Omron CX-Programmer project NewProject (CX-Programmer 9.81)

# PLC masodik: CJ2M CPU32
I/O table (CPU CJ2M-CPU32): rack 0 slot 11 CJ2M-EIP21

## Global symbols (name address type ; comment)
At_entry 2.00 BOOL  ; At entry
At_front 2.06 BOOL  ; At front
At_left_entry 2.08 BOOL  ; At left entry
At_left_exit 2.10 BOOL  ; At left exit
At_load_position 2.04 BOOL  ; At load position
At_right_entry 2.07 BOOL  ; At right entry
At_right_exit 2.09 BOOL  ; At right exit
At_turntable_entry 2.03 BOOL  ; At turntable entry
At_unload_position 2.05 BOOL  ; At unload position
Emergency_stop 2.14 BOOL  ; Emergency stop
Entry_conveyor 3.01 BOOL  ; Entry conveyor
Feeder_conveyor 3.00 BOOL  ; Feeder conveyor
Green_indicator 3.07 BOOL  ; Green indicator
High_box 2.02 BOOL  ; High box
Left_conveyor 3.05 BOOL  ; Left conveyor
Load 3.02 BOOL  ; Load
Low_box 2.01 BOOL  ; Low box
Red_indicator 3.09 BOOL  ; Red indicator
Reset 2.12 BOOL  ; Reset
Reset_light 3.11 BOOL  ; Reset light
Right_conveyor 3.06 BOOL  ; Right conveyor
Start 2.11 BOOL  ; Start
Start_light 3.10 BOOL  ; Start light
Stop 2.13 BOOL  ; Stop
Stop_light 3.12 BOOL  ; Stop light
Turn 3.04 BOOL  ; Turn
Unload 3.03 BOOL  ; Unload
Yellow_indicator 3.08 BOOL  ; Yellow indicator
a_num W350 UINT
b_num W351 UINT
dest W352 UINT
next_prod W200 UINT

## Program NewProgram2 (cyclic task 0)
Local symbols
enable W0.00 BOOL
left_counter W4 UINT
right_counter W5 UINT
stack_length W6 UINT
stack_light UINT
stack_null W0.04 BOOL
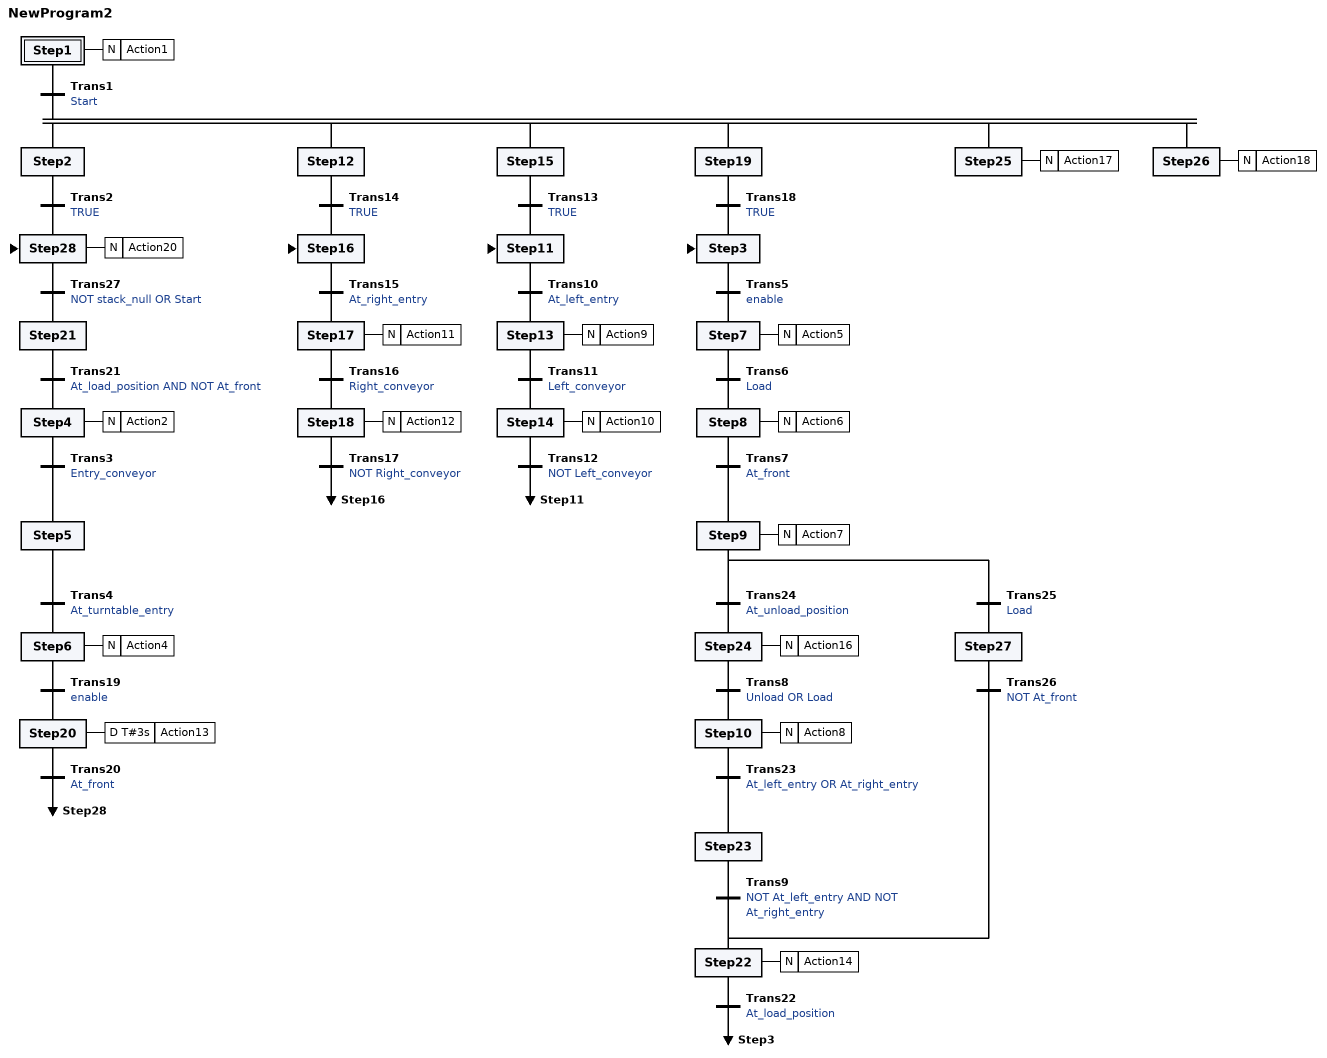
INITIAL_STEP Step1 :
Action1(N) ;
END_STEP
TRANSITION Trans1 FROM Step1 TO (Step2,Step12,Step15,Step19,Step25,Step26)
 := Start;
END_TRANSITION
STEP Step2 :
END_STEP
STEP Step3 :
END_STEP
TRANSITION Trans2 FROM Step2 TO Step28
 := TRUE;
END_TRANSITION
STEP Step4 :
Action2(N) ;
END_STEP
TRANSITION Trans3 FROM Step4 TO Step5
 := Entry_conveyor;
END_TRANSITION
STEP Step5 :
END_STEP
TRANSITION Trans4 FROM Step5 TO Step6
 := At_turntable_entry;
END_TRANSITION
STEP Step6 :
Action4(N) ;
END_STEP
TRANSITION Trans5 FROM Step3 TO Step7
 := enable;
END_TRANSITION
STEP Step7 :
Action5(N) ;
END_STEP
TRANSITION Trans6 FROM Step7 TO Step8
 := Load;
END_TRANSITION
STEP Step8 :
Action6(N) ;
END_STEP
TRANSITION Trans7 FROM Step8 TO Step9
 := At_front;
END_TRANSITION
STEP Step9 :
Action7(N) ;
END_STEP
TRANSITION Trans8 FROM Step24 TO Step10
 := Unload OR Load;
END_TRANSITION
STEP Step11 :
END_STEP
STEP Step12 :
END_STEP
TRANSITION Trans10 FROM Step11 TO Step13
 := At_left_entry;
END_TRANSITION
STEP Step13 :
Action9(N) ;
END_STEP
TRANSITION Trans11 FROM Step13 TO Step14
 := Left_conveyor;
END_TRANSITION
STEP Step14 :
Action10(N) ;
END_STEP
STEP Step10 :
Action8(N) ;
END_STEP
TRANSITION Trans9 FROM Step23 TO Step22
 := NOT At_left_entry AND NOT At_right_entry;
END_TRANSITION
TRANSITION Trans12 FROM Step14 TO Step11
 := NOT Left_conveyor;
END_TRANSITION
STEP Step15 :
END_STEP
TRANSITION Trans13 FROM Step15 TO Step11
 := TRUE;
END_TRANSITION
TRANSITION Trans14 FROM Step12 TO Step16
 := TRUE;
END_TRANSITION
STEP Step16 :
END_STEP
TRANSITION Trans15 FROM Step16 TO Step17
 := At_right_entry;
END_TRANSITION
STEP Step17 :
Action11(N) ;
END_STEP
TRANSITION Trans16 FROM Step17 TO Step18
 := Right_conveyor;
END_TRANSITION
STEP Step18 :
Action12(N) ;
END_STEP
TRANSITION Trans17 FROM Step18 TO Step16
 := NOT Right_conveyor;
END_TRANSITION
STEP Step19 :
END_STEP
TRANSITION Trans18 FROM Step19 TO Step3
 := TRUE;
END_TRANSITION
TRANSITION Trans19 FROM Step6 TO Step20
 := enable;
END_TRANSITION
STEP Step20 :
Action13(D,T#3s) ;
END_STEP
TRANSITION Trans20 FROM Step20 TO Step28
 := At_front;
END_TRANSITION
STEP Step21 :
END_STEP
TRANSITION Trans21 FROM Step21 TO Step4
 := At_load_position AND NOT At_front;
END_TRANSITION
STEP Step22 :
Action14(N) ;
END_STEP
TRANSITION Trans22 FROM Step22 TO Step3
 := At_load_position;
END_TRANSITION
TRANSITION Trans23 FROM Step10 TO Step23
 := At_left_entry OR At_right_entry;
END_TRANSITION
STEP Step23 :
END_STEP
STEP Step24 :
Action16(N) ;
END_STEP
STEP Step25 :
Action17(N) ;
END_STEP
STEP Step26 :
Action18(N) ;
END_STEP
TRANSITION Trans24 (PRIORITY := 1) FROM Step9 TO Step24
 := At_unload_position;
END_TRANSITION
TRANSITION Trans25 (PRIORITY := 2) FROM Step9 TO Step27
 := Load;
END_TRANSITION
STEP Step27 :
END_STEP
TRANSITION Trans26 FROM Step27 TO Step22
 := NOT At_front;
END_TRANSITION
STEP Step28 :
Action20(N) ;
END_STEP
TRANSITION Trans27 FROM Step28 TO Step21
 := NOT stack_null OR Start;
END_TRANSITION

### Action Action1

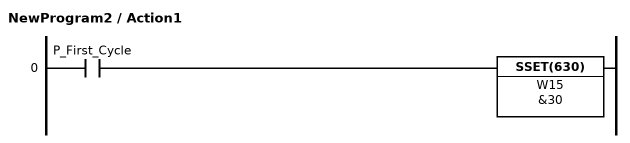
; rung 0
LD P_First_Cycle
SSET(630) W15 &30

### Action Action2

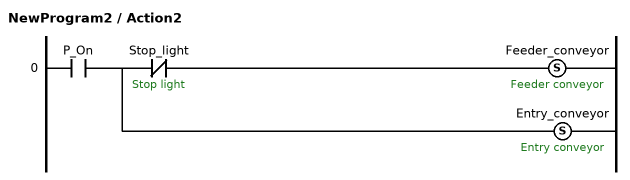
; rung 0
LD P_On
OUT TR0
ANDNOT Stop_light  ; Stop light
SET Feeder_conveyor  ; Feeder conveyor
LD TR0
SET Entry_conveyor  ; Entry conveyor

### Action Action3

### Action Action4

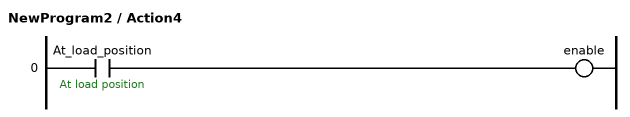
; rung 0
LD At_load_position  ; At load position
OUT enable

### Action Action5

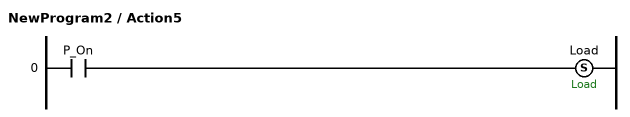
; rung 0
LD P_On
SET Load  ; Load

### Action Action6

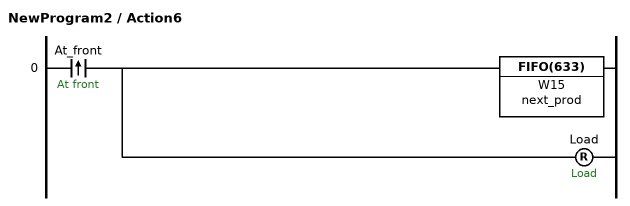
; rung 0
@LD At_front  ; At front
FIFO(633) W15 next_prod
RSET Load  ; Load

### Action Action7

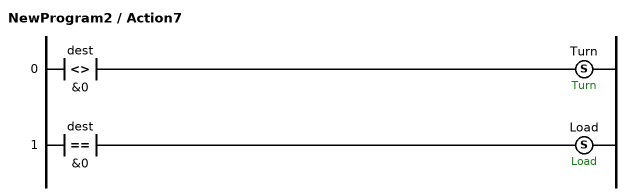
; rung 0
LD<>(305) dest &0
SET Turn  ; Turn
; rung 1
LD=(300) dest &0
SET Load  ; Load

### Action Action8

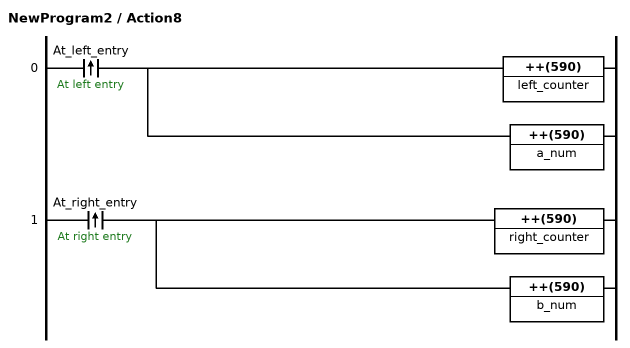
; rung 0
@LD At_left_entry  ; At left entry
++(590) left_counter
++(590) a_num
; rung 1
@LD At_right_entry  ; At right entry
++(590) right_counter
++(590) b_num

### Action Action9

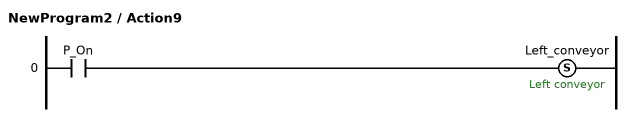
; rung 0
LD P_On
SET Left_conveyor  ; Left conveyor

### Action Action10

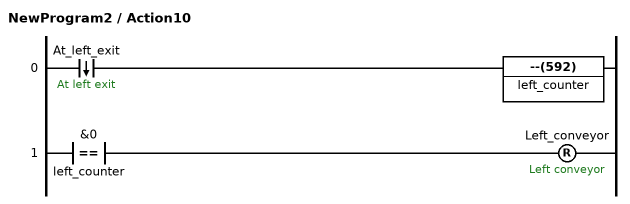
; rung 0
%LD At_left_exit  ; At left exit
--(592) left_counter
; rung 1
LD=(300) &0 left_counter
RSET Left_conveyor  ; Left conveyor

### Action Action11

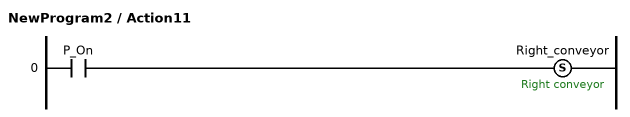
; rung 0
LD P_On
SET Right_conveyor  ; Right conveyor

### Action Action12

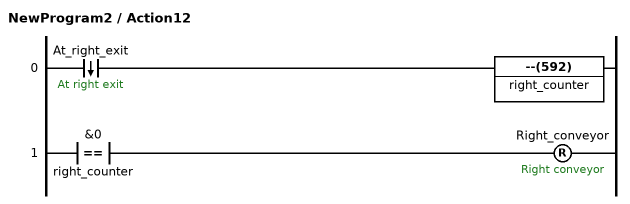
; rung 0
%LD At_right_exit  ; At right exit
--(592) right_counter
; rung 1
LD=(300) &0 right_counter
RSET Right_conveyor  ; Right conveyor

### Action Action13

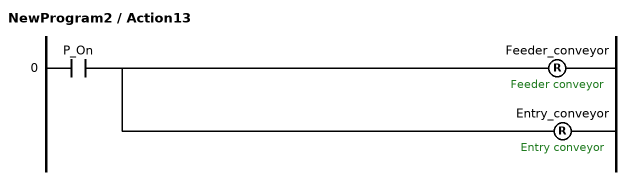
; rung 0
LD P_On
RSET Feeder_conveyor  ; Feeder conveyor
RSET Entry_conveyor  ; Entry conveyor

### Action Action14

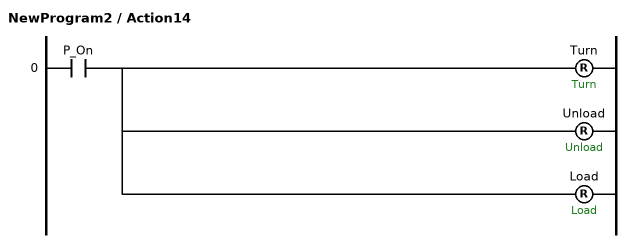
; rung 0
LD P_On
RSET Turn  ; Turn
RSET Unload  ; Unload
RSET Load  ; Load

### Action Action15

### Action Action16

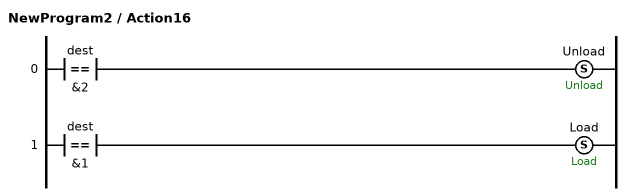
; rung 0
LD=(300) dest &2
SET Unload  ; Unload
; rung 1
LD=(300) dest &1
SET Load  ; Load

### Action Action17

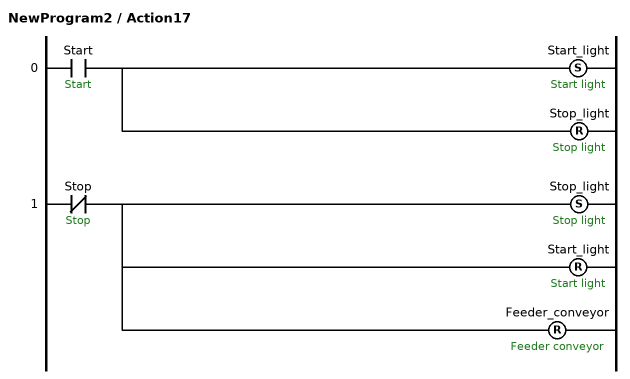
; rung 0
LD Start  ; Start
SET Start_light  ; Start light
RSET Stop_light  ; Stop light
; rung 1
LDNOT Stop  ; Stop
SET Stop_light  ; Stop light
RSET Start_light  ; Start light
RSET Feeder_conveyor  ; Feeder conveyor

### Action Action18

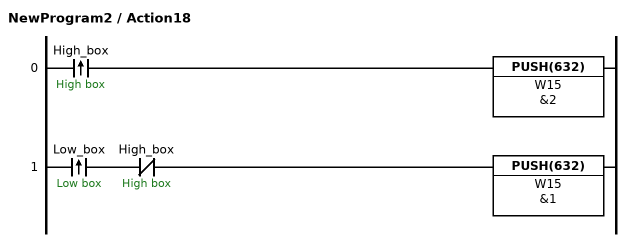
; rung 0
@LD High_box  ; High box
PUSH(632) W15 &2
; rung 1
@LD Low_box  ; Low box
ANDNOT High_box  ; High box
PUSH(632) W15 &1

### Action Action19

### Action Action20

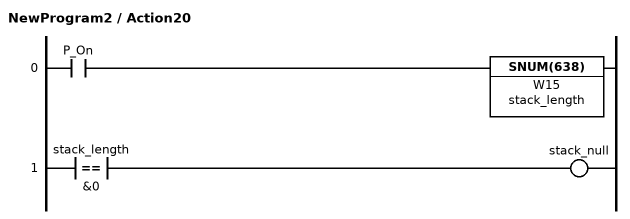
; rung 0
LD P_On
SNUM(638) W15 stack_length
; rung 1
LD=(300) stack_length &0
OUT stack_null

## Program NewProgram3 (cyclic task 1)
Local symbols
a_array W500 UINT[4]
a_comp W0.01 BOOL
b_array W400 UINT[6]
b_comp W0.02 BOOL
IF P_First_Cycle THEN
	a_num := 0;
	b_num := 0;
	a_comp := FALSE;
	b_comp := FALSE;
	
	a_array[0] := 1;
	a_array[1] := 2;
	a_array[2] := 1;
	a_array[3] := 2;
	
	b_array[0] := 1;
	b_array[1] := 1;
	b_array[2] := 1;
	b_array[3] := 2;
	b_array[4] := 2;
	b_array[5] := 2;
END_IF;

IF a_comp AND b_comp THEN
	dest := 0;
ELSIF a_comp AND b_array[b_num] = next_prod THEN
	dest := 2;
ELSIF b_comp AND a_array[a_num] = next_prod THEN
	dest := 1;
ELSIF next_prod = 1 THEN
	IF a_array[a_num] <> 1 AND b_array[b_num] <> 1 THEN
		dest := 0;
	ELSIF a_array[a_num] = 1 AND b_array[b_num] <> 1 THEN
		dest := 1;
	ELSIF a_array[a_num] <> 1 AND b_array[b_num] = 1 THEN
		dest := 2;
	ELSIF a_array[a_num] = 1 AND b_array[b_num] = 1 THEN
		IF a_num > b_num THEN
			dest := 2;
		ELSIF a_num < b_num THEN
			dest := 1;
		ELSE
			dest := 1;
		END_IF;
	END_IF;
ELSIF next_prod = 2 THEN
	IF a_array[a_num] <> 2 AND b_array[b_num] <> 2 THEN
		dest := 0;
	ELSIF a_array[a_num] = 2 AND b_array[b_num] <> 2 THEN
		dest := 1;
	ELSIF a_array[a_num] <> 2 AND b_array[b_num] = 2 THEN
		dest := 2;
	ELSIF a_array[a_num] = 2 AND b_array[b_num] = 2 THEN
		IF a_num > b_num THEN
			dest := 2;
		ELSIF a_num < b_num THEN
			dest := 1;
		ELSE
			dest := 1;
		END_IF;
	END_IF;
END_IF;

## Program NewProgram1 (cyclic task 2)
Local symbols
Emergency_light BOOL
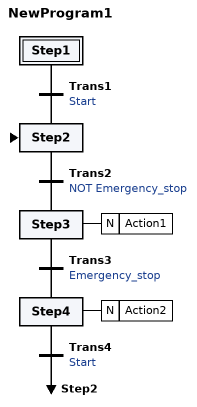
INITIAL_STEP Step1 :
END_STEP
TRANSITION Trans1 FROM Step1 TO Step2
 := Start;
END_TRANSITION
STEP Step2 :
END_STEP
TRANSITION Trans2 FROM Step2 TO Step3
 := NOT Emergency_stop;
END_TRANSITION
STEP Step3 :
Action1(N) ;
END_STEP
TRANSITION Trans3 FROM Step3 TO Step4
 := Emergency_stop;
END_TRANSITION
STEP Step4 :
Action2(N) ;
END_STEP
TRANSITION Trans4 FROM Step4 TO Step2
 := Start;
END_TRANSITION

### Action Action1

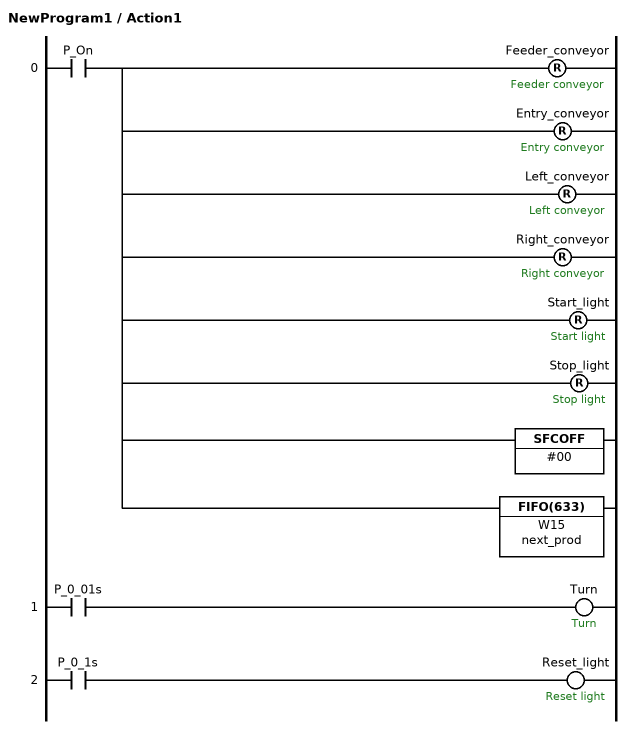
; rung 0
LD P_On
RSET Feeder_conveyor  ; Feeder conveyor
RSET Entry_conveyor  ; Entry conveyor
RSET Left_conveyor  ; Left conveyor
RSET Right_conveyor  ; Right conveyor
RSET Start_light  ; Start light
RSET Stop_light  ; Stop light
SFCOFF #00
FIFO(633) W15 next_prod
; rung 1
LD P_0_01s
OUT Turn  ; Turn
; rung 2
LD P_0_1s
OUT Reset_light  ; Reset light

### Action Action2

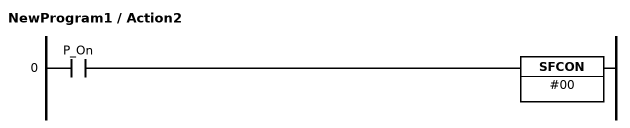
; rung 0
LD P_On
SFCON #00